  def clear_poses():
      pose = create_transition_pose()
      pose_start = create_transition_pose()
      pose_help = create_transition_pose()
      pose_target = create_transition_pose()
  end

  def do_transition(reference_pose=p[0,0,0,0,0,0], mode=2, keep_rxry=False, a=1.4, v=1.05, r=0.100):
      # the robot will evaluate the current and target workarea
      # after that, the robot will move between the workareas automatically.
      # parameters:
      # reference_pose:   a pose/frame were the robot should work next. If nothing is given, base frame will be used as target
      # keep_rxry:        if true, the robot will keep the orientation of the tool during the movement

      ################# checking #################
      clear_poses()
      workarea_current = check_workarea(get_actual_tcp_pose())    # between 0 and the amount of defined workareas
      workarea_new = check_workarea(reference_pose)               # between 0 and the amount of defined workareas
      reverse_rotation = False

      if (workarea_current != 0 and workarea_new != 0 and workarea_current != workarea_new) or (reference_pose == p[0,0,0,0,0,0]):
          ################# get axisvalues #################
          if (mode == 1):
              pose_start = get_transition_pose_by_workarea(workarea_current)
              pose_target = get_transition_pose_by_workarea(workarea_new)
          elif (mode == 2):
              pose_start = get_transition_pose_by_reference_pose(get_actual_tcp_pose(), RADIUS_TRANSITION_POSES, keep_rxry)
              pose_target = get_transition_pose_by_reference_pose(reference_pose, RADIUS_TRANSITION_POSES, keep_rxry)

          end
          # if (pose_start.crt[1] < 0 and pose_target.crt[1] > 0) or (pose_start.crt[1] > 0 and pose_target.crt[1] < 0):
          #     pose_help = get_transition_pose_by_reference_pose(pose_start.crt, RADIUS_HELPER_POSES)
          # end
          textmsg("Cartesian pose start: ", to_str(pose_start.crt))
          textmsg("Joints pose start: ", to_str(pose_start.jnt))
          textmsg("Qnear pose start: ", to_str(pose_start.q))
          textmsg("Cartesian pose target: ", to_str(pose_target.crt))
          textmsg("Joints pose target: ", to_str(pose_target.jnt))
          textmsg("Qnear pose target: ", to_str(pose_target.q))

          ################# movements #################
          if (pose_help.jnt != [0,0,0,0,0,0]):
              if point_dist(get_actual_tcp_pose(), pose_start.crt) > r and point_dist(pose_start.crt, pose_help.crt) > r:
                  movej(pose_start.jnt, a=a, v=v, r=r)
                  if (point_dist(pose_start.crt, pose_help.crt) > r) and (point_dist(pose_target.crt, pose_help.crt) > r):
                      movej(pose_help.jnt, a=a, v=v, r=r)
                  end
              end
          else:
              if point_dist(get_actual_tcp_pose(), pose_start.crt) > r and point_dist(pose_start.crt, pose_target.crt) > r:
                  movej(pose_start.jnt, a=a, v=v, r=r)
              end
          end
          movej(pose_target.jnt, a=a, v=v)

          ################# checking #################
          workarea_current = check_workarea(get_actual_tcp_pose())    # between 0 and the amount of defined workareas
      else:
          # define error or warning
      end
  end


  # Erläuterung
  # für start wird die aktuelle Position übergeben
  # davon wird die Position für start berechnet. Bei der Orientierung wird entweder nur Rz genommen oder alles bei keep_rxry
  $ 11 "Script: SCRIPT Logs V1.2.script"
  current_state_log = ""
  current_process_log = ""
  current_step_log = ""
  current_warning_log = ""
  current_error_log = ""
  current_hatch_log = ""
  current_centrifuge_log = ""
  current_message_log = "placeholderstring"
  LogLevel=struct(NONE=0, INFO=1, PROCESS=2, WARNING=3, ERROR=4)
  LOGLEVEL=LogLevel.INFO

  def log_message(prefix="", newlog=current_message_log):
      # generates a log message every time its useful
      if (current_message_log != newlog and newlog != ""):
          textmsg(str_cat(prefix, to_str(newlog)))
          current_message_log = to_str(newlog)
      end
  end

  def log_state(newlog):
      # generates a log message every time its useful
      if (current_state_log != newlog and newlog != ""):
          textmsg(str_cat("Machine: ", to_str(newlog)))
          current_state_log = to_str(newlog)
      end
  end

  def log_process(newlog):
      # generates a log message every time its useful
      if (current_process_log != newlog and newlog != ""):
          textmsg(str_cat("Process: ", to_str(newlog)))
          current_process_log = to_str(newlog)
      end
  end

  def log_step(newlog):
      # generates a log message every time its useful
      if (current_step_log != newlog and newlog != ""):
          textmsg(str_cat("Step: ", to_str(newlog)))
          current_step_log = to_str(newlog)
      end
  end

  def log_info(newlog):
      # generates a log message if log level is Info or lower
      if (newlog != "" and LOGLEVEL <= LogLevel.INFO):
          textmsg(str_cat("INFO: ", newlog))
      end
  end

  def log_warning(newlog):
      # generates a log message every time its useful
      if (current_warning_log != newlog and newlog != ""):
          textmsg(str_cat("WARNING: ", to_str(newlog)))
          current_warning_log = to_str(newlog)
      end
  end

  def log_error(newlog):
      # generates a log message every time its useful
      if (current_error_log != newlog and newlog != ""):
          textmsg(str_cat("ERROR: ", to_str(newlog)))
          current_error_log = to_str(newlog)
      end
  end

  def log_hatch_state(newlog):
      # generates a log message every time its useful
      if (current_hatch_log != to_str(newlog) and to_str(newlog) != ""):
          textmsg(str_cat("Hatch_state: ", to_str(newlog)))
          current_hatch_log = to_str(newlog)
      end
  end

  def log_centrifuge_state(newlog):
      # generates a log message every time its useful
      if (current_centrifuge_log != to_str(newlog) and to_str(newlog) != ""):
          textmsg(str_cat("Centrifuge_state: ", to_str(newlog)))
          current_centrifuge_log = to_str(newlog)
      end
  end
  $ 12 "Script: SCRIPT Statistics V1.1.script"
  #*****************************************************
  # customer          :   tbd
  # project name      :   tbd
  #****************************************************
  # controller        :
  # software          :
  #****************************************************
  # author            :   P. Koehnke (+49 1628859904; p.koehnke@unitedrobotics.group)
  # Copyright (c)     :   United Robotics Group Health and Food GmbH
  #                       An der Riede 2
  #                       28816 Stuhr
  #                       Germany
  #****************************************************
  # description       :   statistics script, which tracks the times in different PackML states and let you count objects
  # version:      	:   1.0
  # created           :   20.11.2023
  # updated           :
  #****************************************************
  # modifications     :
  #
  # date              :
  # name              :
  # reason            :
  #****************************************************

  # to save the times persistently, these variables must be defined in the installation file of the robot

  # ===== object counters =====
  def count_up(counters, idx, by):
      counters[idx] = counters[idx] + by
      return counters
  end

  def count_total(counters):
      local i = 0
      local total = 0
      while (i<length(counters)):
          total = total + counters[i]
          i = i + 1
      end
      return total
  end
  # ==========

  # ===== Times =====
  thread Pml_Timer_Thread():
      # STATE_Times is a list of all time values in seconds
      while (True):
          STATE_Times[STATE-1] = STATE_Times[STATE-1] + get_steptime()
          sync()
      end
  end

  thread_timer_handler = run Pml_Timer_Thread()

  def get_time(timer, format="dd/hh/mm/ss"):
      # give the time in seconds
      # the function will return the given time as string in the predefined format
      local days = floor(timer/86400)
      local hours = floor((timer%86400)/3600)
      local minutes = floor((timer%3600)/60)
      local seconds = floor(timer%60)
      return str_cat(str_cat(str_cat(str_cat(str_cat(str_cat(to_str(days), "/"), to_str(hours)), "/"), to_str(minutes)), "/"), to_str(seconds))
  end

  def set_timer(time, format="dd/hh/mm/ss"):
      # give the time as string
      # the function will return the corresponding seconds summed up
      local days_idx = str_find(time, "/", 0)
      local hours_idx = str_find(time, "/", days_idx+1)
      local minutes_idx = str_find(time, "/", hours_idx+1)
      local days = to_num(str_sub(time, 0, days_idx))
      local hours = to_num(str_sub(time, days_idx+1, hours_idx-days_idx-1))
      local minutes = to_num(str_sub(time, hours_idx+1, minutes_idx-hours_idx-1))
      local seconds = to_num(str_sub(time, minutes_idx+1, length(time)-minutes_idx))
      return (days*86400 + hours*3600 + minutes*60 + seconds)
  end
  $ 13 "Script: SCRIPT Vision Config V0.2.script"
  CAM_LM = struct(id=0, type="", size=0, related_itm=0, capture_relation="")
  global CAM_Result = make_list(0, 0, 50)

  def create_landmark(id=0, type="", size=0, related_itm=0, capture_relation=""):
      return struct(id=id, type=type, size=size, related_itm=related_itm, capture_relation=capture_relation)
  end


  CAM_LMs = [
    create_landmark(id=1, type="aruco_7x7", size=0.1, related_itm=1, capture_relation="front_right"),
    create_landmark(id=4, type="aruco_7x7", size=0.1, related_itm=2, capture_relation="straight_left"),
    create_landmark(id=3, type="aruco_7x7", size=0.1, related_itm=2, capture_relation="straight_left"),
    create_landmark(id=8, type="aruco_7x7", size=0.1, related_itm=2, capture_relation="right"),
    create_landmark(id=5, type="aruco_7x7", size=0.1, related_itm=5, capture_relation="left"),
    create_landmark(id=6, type="aruco_7x7", size=0.1, related_itm=2, capture_relation="straight_left")
  ]

  CAM_Capture_Poses = struct(
    front_left = p[0.350,-0.330,0.500,0.353,-0.323,-1.458],
    left = p[0.350,0.000,0.500,0.353,-0.323,-1.458],
    back_left = p[0.350,0.220,0.500,0.353,-0.323,-1.458],
    back_right = p[-0.350,0.000,0.500,0.579,0.240,0.760],
    right = p[-0.350,-0.300,0.500,0.206,0.206,1.561],
    front_right = p[-0.350,-0.400,0.500,0.242,0.903,2.480],
    straight_left = p[0.375,-0.000,0.500,0.815,-0.815,-1.412],
    front = p[0,0,0,0,0,0]
  )

  def get_capture_pose(lm):
      if (lm.capture_relation == "front_left"):
          return CAM_Capture_Poses.front_left
      elif (lm.capture_relation == "left"):
          return CAM_Capture_Poses.left
      elif (lm.capture_relation == "back_left"):
          return CAM_Capture_Poses.back_left
      elif (lm.capture_relation == "back_right"):
          return CAM_Capture_Poses.back_right
      elif (lm.capture_relation == "right"):
          return CAM_Capture_Poses.right
      elif (lm.capture_relation == "straight_left"):
         return CAM_Capture_Poses.straight_left
      else:
          # error
          return get_actual_tcp_pose()
      end
  end
  $ 14 "Script: SCRIPT uLM Factory.script"
  # ############### SCRIPT uLM Factory ##################
  # *****************************************************
  # Customer          :   URG
  # Product Name      :   uLabMobile
  # ****************************************************
  # Controller/Robot  :   UR5e
  # Software          :   URSCRIPT
  # Dependencies      :   Defines Script but mainly independend
  # How To            :   is used by projectconfig to create list of structs full of projectrelated information which are used across the scripts
  # ****************************************************
  # Author            :   D.Kreugel
  # Copyright (c)     :   United Robotics Group Health and Food GmbH
  #                       An der Riede 2
  #                       28816 Stuhr
  #                       Germany
  # ****************************************************
  # Description       :   definition of the datastructures used by the uLM, gives functionality to create a predefined datastructure, is assigned to a global list in projectconfig
  # Version           :   0.2
  # Created           :   18.07.2024
  # Updated           :
  # ****************************************************
  # Modifications     :
  #
  # Date              :
  # Name              :
  # Reason            :
  # ****************************************************
  # TODO              : cleanup useless info and add all other factorys from the other scripts here to have one place to search for such things, documentation

  # DO NOT TOUCH THE DATASTRUCTURES IF YOU DON'T KNOW WHAT YOU DO!
  MAX_ACTIONS=6
  POS_Z=p[0,0,0,0,0,0]
  def create_pattern(id=0, name="", pattern_width=[0, 0], pattern_size=[0, 0], blocked=[-1, -1, -1], direction="X", transpose=False, invert=False, description="default"):
      return struct(
          id = id,
          name = name,
          pattern_width = pattern_width,
          pattern_size = pattern_size,
          blocked = blocked,
          direction = direction,
          transpose = transpose,
          invert = invert,
          description = description
      )
  end

  # item model stores frame related inner and outer patterns
  def create_item_model(inner="", outer="", description="default"):
      return struct(
          inner = inner,
          outer = outer,
          description = description
          )
  end

  # creates a fixed length list cause structs cannot deal with dynamic lists at the moment and an item can have different amount of actions assigned to it
  def create_action_list(values):
      local list = make_list(MAX_ACTIONS, 0, MAX_ACTIONS+1)
      local i = 0
      while (i < values.length()):
          list[i] = values[i]
          i = i + 1
      end
      return list
  end

  def create_item(id=0, ls_item="default", frame=p[0,0,0,0,0,0], actionlist=create_action_list([]), item_model=create_item_model(), lm_id=0, description="default"):
      return struct(
          id = id,
          ls_item = ls_item,
          frame = frame,
          actionlist = create_action_list(actionlist),
          item_model = item_model,
          lm_id = lm_id,
          description = description
      )
  end

  def create_object(id=0, obj_name=0, height=0, width=0, obj_type = 0, description="default"):
      return struct(
          id = id,
          obj_name = obj_name,
          obj_type = obj_type,
          height = height,
          width = width,
          description = description
      )
  end
  # extends object type by sample related information
  def create_sample(obj_id=0, cap_diameter=0, raw_diameter=0, color="", material="", description=""):
      return struct(
      obj_id = obj_id,
      cap_diameter = cap_diameter,
      raw_diameter = raw_diameter,
      color = color,
      material = material,
      description = description)
  end

  # create gripper configs
  def create_gripper_config(gripper_offset=struct(prepick=2, pick=0, place=2), force=0, speed=0, validation=0, object=create_object()):
      gripper_offset.prepick = object.width+gripper_offset.prepick
      gripper_offset.place = object.width+gripper_offset.place
      return struct(
          object = object.obj_name,
          force = force,
          speed = speed,
          validation = validation,
          width = gripper_offset
      )
  end

  def create_manipulator_command(id="", item="", action=0, jig_nbr=-1, obj_nbr=-1, object_type=-1, error_id=0, data=""):
      return struct(
          id = id,
          device = Device.MANIPULATOR,
          item = item,
          action = action,
          jig_nbr = jig_nbr,
          obj_nbr = obj_nbr,
          object_type = object_type,
          error_id = error_id,
          data = data
      )
  end

  def create_amr_command(id="", item="", action=0, target=0, error_id=0, data=""):
      return struct(
          id = id,
          device = Device.AMR,
          item = item,
          action = action,
          target = target,
          error_id = error_id,
          data = data
      )
  end

  def create_camera_command(id="", item="", action=0, attempt=0, error_id=0, data=""):
      return struct(
          id = id,
          device = Device.CAMERA,
          item = item,
          action = action,
          attempt = attempt,
          error_id = error_id,
          data = data
      )
  end

  # Function to create a new  vision struct to assign workspace and skill to an item or a selection
  def create_vision_config(workspace_id="", skill_id="", item_id=-1, target_origin=p[0,0,0,0,0,0], description="default"):
      return struct(
          workspace_id = workspace_id,
          skill_id = skill_id,
          item_id = item_id,
          target_origin = target_origin,
          description = description)
  end

  # extents the vision config by the inspect configuration, this info will be called in the action inspect only
  # item_id is the reference to the item
  # dx is the distance in x direction for one position to the next in the inspection rack
  # dy is the distance in y direction for one position to the next in the inspection rack
  # target origin is the origin coordinate of the first position in the inspectionrack from where the calculation starts
  def create_inspect_config(item_id=0, dx=0, dy=0, target_origin=p[0,0,0,0,0,0], rack_size=[0,0], description="default"):
      return struct(
      item_id = item_id,
      dx = dx,
      dy = dy,
      target_origin = target_origin,
      rack_size = rack_size,
      description = description
      )
  end
   # Function to create a new landmark struct that contains all lm related configurationparameters and will be assigned via item_id
  #def create_landmark(lm_id=0, marker_id=-1, marker_size=0.1, marker_type="aruco_7x7", capture_pos=p[0,0,0,0,0,0], init_frame=p[0,0,0,0,0,0], search_offset=[0,0,0], actual_frame=p[0,0,0,0,0,0], description=""):
    ##  return struct(
     #     lm_id = lm_id,
     #     marker_id = marker_id,
       #   marker_size = marker_size,
    ##      marker_type = marker_type,
    #      capture_pos = capture_pos,
    #      init_frame = init_frame,
    #      search_offset = search_offset,
    #      actual_frame = actual_frame,
  #        description = description)
  #end

  def create_movement(id=0, actionlist=create_action_list([]), hh_approach=POS_Z, h_approach=POS_Z, approach=POS_Z, h_target=POS_Z, target=POS_Z, retract=POS_Z, h_retract=POS_Z, hh_retract=POS_Z, h_frame=POS_Z, frame=POS_Z, speed=1, acceleration=1, description="default"):
  return struct(
      id = id,
      actionlist = actionlist,
      hh_approach = hh_approach,
      h_approach = h_approach,
      approach = approach,
      h_target = h_target,
      target = target,
      retract = retract,
      h_retract = h_retract,
      hh_retract = hh_retract,
      h_frame = h_frame,
      frame = frame,
      speed = speed,
      acceleration = acceleration,
      description = description
  )
  end






  $ 15 "Script: SCRIPT uLM Defines v0.2.script"
  ############# SCRIPT uLM Defines ###############
  #*****************************************************
  # Customer          :   URG
  # Product Name      :   uLabMobile
  #****************************************************
  # Controller/Robot  :   UR5e
  # Software          :   5.17
  # Dependencies      :   Factory Script, Logs Script
  # How To            :   Define Constants depending on the Project, don't go to big in Listsize as it will exceed the URScript limits
  #****************************************************
  # Author            :   D.Kreugel
  # Copyright (c)     :   United Robotics Group Health and Food GmbH
  #                       An der Riede 2
  #                       28816 Stuhr
  #                       Germany
  #****************************************************
  # Description       :   Defines all Enums and Global reachable Varibles/Datastructures
  # Version           :   0.2
  # Created           :   18.07.2024
  # Updated           :
  #****************************************************
  # Modifications     :
  #
  # Date              :
  # Name              :
  # Reason            :
  #****************************************************
  # TODO find better place for the Search Funktions for the Object Lists, documentation


  POS_Z = p[0,0,0,0,0,0]

  # DEFAULTS ROBOT MOVEMENTS
  DEFAULT = struct(SPEED=0.8, ACCELERATION=0.6)

  # ENUMS
  Objects = struct(NONE=0, CC_SAMPLE=1, CC_RACK=2, COAG_SAMPLE=3, COAG_RACK=4, HEMA_SAMPLE=5, HEMA_RACK=6, INPUT_RACK=7, CF_RACK=8, ANY_SAMPLE=9, ANY_RACK=10, TARA_SAMPLE=11, BUTTON=12, XN550_DRAWER=13, COBAS_RACK=14)
  ObjectType = struct(NONE=0,SAMPLE=1,RACK=2, BUTTON=3, DRAWER=4)

  ActionManipulator = struct(NONE=0, PICK=1, PLACE=2, DECAP=12, PUSH=3, RELEASE=21, GRASP=20, MOVE_TO=19, DRAWER_OPEN=51, DRAWER_CLOSE=52)
  ActionAMR = struct(NONE=0, LOAD_MISSION=31, START_MISSION=32, NAVIGATE=33, ACKNOWLEDGE=34, READ=35)
  ActionCamera = struct(NONE=0, INSPECT=16, DETECT=15, DETECT_OBJECTS=17)
  Device = struct(MANIPULATOR=1, AMR=2, CAMERA=3)
  Patterns = struct(NONE="NONE", TARA="TARA", CENTRIFUGE="CENTRIFUGE",CENTRIFUGE_MAGAZINE="CENTRIFUGE_MAGAZINE",SYSMEX_XN550="SYSMEX_XN550",COBAS="COBAS",COBAS_MAGAZINE="COBAS_MAGAZINE",INPUT="INPUT",NOK="NOK",DRAWER_XN550="DRAWER_XN550",ARCHIVE="ARCHIVE")
  CommandStatus = struct(EXECUTED=0, UNFINISHED=1)

  # Constants
  MAX_CAPTURE_ATTEMPTS = 8
  # Maximum Size of the Datastructures
  MAX_ITEM_OBJ = 40
  MAX_GRIPPER_OBJ = 10
  MAX_LANDMARK_OBJ = 10
  MAX_PATTERN_OBJ = 30
  MAX_ITEM_MODEL_OBJ = 20
  MAX_VISION_CONFIG_OBJ = 10
  MAX_CAPTURE_RESULTS = 55
  MAX_MOVEMENT_OBJ = 50

  CON=False

  # for Marburg Approach
  LAST_CAPTURE = make_list(0, "", MAX_CAPTURE_RESULTS)

  # Initialize the Datastructures in order to store related Data and use them in structs without length issues

  OBJECT_MAP = make_list(0 ,create_object(), MAX_ITEM_OBJ)
  ITEM_MAP = make_list(0, create_item(), MAX_ITEM_OBJ)
  ITEM_MODEL_MAP = make_list(0, create_pattern(), MAX_ITEM_MODEL_OBJ)
  GRIPPER_CONFIG_MAP = make_list(0, create_gripper_config(), MAX_PATTERN_OBJ)
  VISION_CONFIG_MAP = make_list(0, create_vision_config(), MAX_VISION_CONFIG_OBJ)
  INSPECT_CONFIG_MAP = make_list(0, create_inspect_config(), MAX_VISION_CONFIG_OBJ)
  LANDMARK_MAP = make_list(0, create_landmark(), MAX_LANDMARK_OBJ)
  MOVEMENT_MAP = make_list(0, create_movement(), MAX_MOVEMENT_OBJ)

  OBJECT_REFERENCE_HEIGHT = 81


  # functions to search in the datastructures which are defined in the factories

  ################# MOVEMENT ###############

  def find_movement_by_frame_and_action(frame,action):
      local i = 0
      local ii = 0
      while (i < MOVEMENT_MAP.length()):
          if (MOVEMENT_MAP[i].frame == frame):
              while(ii < MOVEMENT_MAP[i].actionlist.length()):
                  if (MOVEMENT_MAP[i].actionlist[ii] == action):
                      log_info("Movement found: [" + to_str(MOVEMENT_MAP[i].description) + "]")
                      return MOVEMENT_MAP[i]
                  end
                  ii = ii + 1
              end
              ii = 0
          end
          i = i + 1
      end
      log_warning("no movement found for frame: [" + to_str(frame) + "]")
      return create_movement(frame=frame)  # Return default pattern if not found
  end

  def find_item_by_lsitem_and_action(ls_item, action):
      local i = 0
      while (i < ITEM_MAP.length()):
          if (ITEM_MAP[i].ls_item == ls_item):
              local ii = 0
              while (ii < ITEM_MAP[i].actionlist.length()):
                  if (ITEM_MAP[i].actionlist[ii] == action):
                      log_info("Item found: [" + to_str(ITEM_MAP[i].description) + "]")
                      return ITEM_MAP[i]
                  end
                  ii = ii + 1
              end
          end
          i = i + 1
      end
      log_warning("Item not found for station[" + to_str(ls_item) + "] and action[" + to_str(action) + "]")
      return create_item()  # Return default item if not found
  end
  ################# PATTERN ###################

  def find_pattern_by_name(name):
      local i = 0
      while (i < ITEM_MODEL_MAP.length()):
          if (ITEM_MODEL_MAP[i].name == name):
              log_info("Item Model found: [" + to_str(ITEM_MODEL_MAP[i].description) + "]")
              return ITEM_MODEL_MAP[i]
          end
          i = i + 1
      end
      log_warning("Item Model not found for name[" + to_str(name) + "]")
      return create_pattern()  # Return default pattern if not found
  end

  def is_in_list(list,val):
      local i = 0
      while(i<list.length()):
          if(list[i]==val):
              return True
          end
          i=i+1
      end
      return False
  end

  def get_next_valid_patternslot(item_model, counter):
      local i = 0
      local temp = 0
      local max_slots = item_model.pattern_size[0] * item_model.pattern_size[1]
      log_info("blocked positions:" + to_str(item_model.blocked) + "| current pos: " + to_str(counter))
      while (i < item_model.blocked.length()):
          if(item_model.blocked[i] <= counter and item_model.blocked[i] != -1):
              temp = temp + 1
          end
          i = i + 1
      end

      if(is_in_list(item_model.blocked,counter+temp)):
          while(is_in_list(item_model.blocked,counter+temp)):
              temp=temp+1
          end
      end
      log_info("changed position in rack to nbr:" + to_str(counter+temp))

      return counter+temp

  end

  ################# OBJECT ###################

  # def find_object_by_material(material):
  #   local i = 0
  #   log_info("Trying to find object by color:", to_str(material))
  #   while (i < OBJECT_MAP.length()):
  #       if (OBJECT_MAP[i].material == material):
  #           log_info("Object model found:", to_str(OBJECT_MAP[i]))
  #           return OBJECT_MAP[i]
  #       end
  #       i = i + 1
  #   end
  #   return OBJ_DEFAULT  # Return default pattern if not found
  # end

  def find_object_by_objectname(objectname):
      local i = 0
      #log_info("Trying to find object by color:", to_str(objectname))
      while (i < OBJECT_MAP.length()):
          if (OBJECT_MAP[i].obj_name == objectname):
              log_info("Object Model found: [" + to_str(OBJECT_MAP[i].description) + "]")
              return OBJECT_MAP[i]
          end
          i = i + 1
      end
      log_warning("no Object Model found for objectname:[" + to_str(objectname) + "]")
      return create_object()
  end

  def find_smallest_object():
      local i = 0
      local min_size = OBJECT_MAP[0].height
      #log_info("Trying to find object by color:", to_str(objectname))
      while (i < OBJECT_MAP.length()):
          if (OBJECT_MAP[i].height <= min_size and OBJECT_MAP[i].height != 0):
              log_info("smaller object found: [" + to_str(OBJECT_MAP[i].description) + "]")
              min_size = OBJECT_MAP[i].height
          end
          i = i + 1
      end
      return min_size
  end

  def find_gripper_config_by_objectname(objectname):
  local i = 0
  while (i < GRIPPER_CONFIG_MAP.length()):
      #log_info("gripper config:",to_str(GRIPPER_CONFIG_MAP[i]))
      if (GRIPPER_CONFIG_MAP[i].object == objectname):
          log_info("found gripper parameters [" + to_str(GRIPPER_CONFIG_MAP[i]) + "]")
          return GRIPPER_CONFIG_MAP[i]
      end
      i = i + 1
  end

  log_warning("no gripper parameters found for object type: " + to_str(objectname))
  return create_gripper_config()
  end
  # Function to find a landmark by item
  def find_landmark_by_id(lm_id):
      local i = 0
      while i < LANDMARK_MAP.length():
          if LANDMARK_MAP[i].lm_id == lm_id:
              log_info("found landmark with id(" + to_str(lm_id) + "): [" + to_str(LANDMARK_MAP[i].description) + "]")
              return LANDMARK_MAP[i]
          end
          i = i + 1
      end
      log_warning("landmark not found for lm_id [" + to_str(lm_id) + "]")
      return create_landmark()
  end
  # Function to find a landmark by item
  def find_landmark_by_capture_pos(capture_pos):
      local i = 0
      while i < LANDMARK_MAP.length():
          if LANDMARK_MAP[i].capture_pos == capture_pos:
              log_info("found landmark by capture_pos [" + to_str(LANDMARK_MAP[i].description) + "]")
              return LANDMARK_MAP[i]
          end
          i = i + 1
      end
      log_warning("Landmark not found for capture_pos: [" + to_str(capture_pos) + "]")
      return create_landmark()
  end

  def update_landmark_by_capture_pos(capture_pos, lm_pos):
      local i = 0
      while i < LANDMARK_MAP.length():
          if LANDMARK_MAP[i].capture_pos == capture_pos:
              log_info("updated landmark from [" + to_str(LANDMARK_MAP[i].description) + "]")
              LANDMARK_MAP[i].actual_frame = lm_pos
              return True
          end
          i = i + 1
      end
      log_warning("Landmark not found for capture_pos: [" + to_str(capture_pos) + "]")
      return False
  end

  def update_landmark_by_id(lm_id,lm_pos):
      local i = 0
      while i < LANDMARK_MAP.length():
          if LANDMARK_MAP[i].lm_id == lm_id:
              log_info("updated landmark.actual_frame from [" + to_str(LANDMARK_MAP[i].description + "]"))
              LANDMARK_MAP[i].actual_frame = lm_pos
              return True
          end
          i = i + 1
      end
      log_warning("Landmark not found for lm_id " + to_str(lm_id))
      return False
  end

  def find_vision_config_by_frame(frame):
      local i = 0
      while i < VISION_CONFIG_MAP.length():
          if VISION_CONFIG_MAP[i].capture_pos == frame:
              log_info("Vision Config found: [" + to_str(VISION_CONFIG_MAP[i].description) + "]")
              return VISION_CONFIG_MAP[i]
          end
          i = i + 1
      end
      log_info("Vision Config not found for frame: " + to_str(frame))
      return create_vision_config()
  end

  def find_vision_config_by_itemid(id):
      local i = 0
      while i < VISION_CONFIG_MAP.length():
          if VISION_CONFIG_MAP[i].item_id == id:
              log_info("Vision Config found: [" + to_str(VISION_CONFIG_MAP[i].description) + "]")
              return VISION_CONFIG_MAP[i]
          end
          i = i + 1
      end
      log_info("Vision Config not found for item: " + to_str(id))
      return create_vision_config()
  end

  def find_inspect_config_by_itemid(id):
      local i = 0
      while i < INSPECT_CONFIG_MAP.length():
          if INSPECT_CONFIG_MAP[i].item_id == id:
              log_info("Inspect Config found: [" + to_str(INSPECT_CONFIG_MAP[i].description) + "]")
              return INSPECT_CONFIG_MAP[i]
          end
          i = i + 1
      end
      log_info("Inspect Config not found for item: " + to_str(id))
      return create_inspect_config()
  end
  $ 16 "Script: SCRIPT Device Robotiq Greifer v0.2.script"
  # ############ SCRIPT Device Robotiq Greifer ###############
  # **********************************************************
  # Customer          :   URG
  # Product Name      :   uLabMobile
  # **********************************************************
  # Controller/Robot  :   UR5e
  # Software          :   5.17
  # Dependencies      :   Logs Script, Robotiq Gripper and Gripper Datastructure for args (Factory Script), URCAP Robotiq
  # **********************************************************
  # Author            :   D.Kreugel, P.Köhnke
  # Copyright (c)     :   United Robotics Group Health and Food GmbH
  #                       An der Riede 2
  #                       28816 Stuhr
  #                       Germany
  # *********************************************************
  # Description       :   Gripper Robotiq Device Interface for Robotiq E-Hand Gripper
  # Version           :   0.2
  # Created           :   18.07.2024
  # Updated           :
  # *********************************************************
  # Modifications     :
  #
  # Date              :
  # Name              :
  # Reason            :
  # *********************************************************
  # TODO              :   documentation

  # RobotiQ Gripper
  ROBOTIQ_GRP_CLOSE = 0
  ROBOTIQ_GRP_OPEN = 40

  # #############FORCEMODE###############
  ROBOTIQ_GRP_FORCE = struct(FULL=100, HALF=50, LOW=25, NONE=0)

  # #############SPEED###################
  ROBOTIQ_GRP_SPEED = struct(FAST=100, MEDIUM=50, SLOW=20)

  # ############VALIDATION###############
  ROBOTIQ_GRP_VALIDATION = struct(ON=1, OFF=0, SKIP=-1)

  # struct(prepick=0, pick=0, place=0, force=0, speed=0, validation=0, object_type=0, description="default")
  def gripper_robotiq_activate():
      return rq_activate_and_wait()
  end

  def gripper_robotiq_reset_and_activate():
      return rq_reset_and_activate()
      #return rq_reset()
  end

  def gripper_robotiq_is_activated():
      return rq_is_gripper_activated()
  end

  def gripper_robotiq_get_current_pos_mm():
      return rq_current_pos_mm()
  end
  # Function to check if the RobotiQ gripper has an object
  def gripper_robotiq_has_object():
      result = rq_is_object_detected()
      if result == False:
          log_error("No object detected by the gripper")
      end
      return result
  end

  def gripper_robotiq_move_to_mm(mm):
      if(gripper_robotiq_is_activated() == False):
          gripper_robotiq_activate()
      end
      return rq_move_and_wait_mm(mm)
  end

  def gripper_robotiq_close():
      if(gripper_robotiq_is_activated() == False):
          gripper_robotiq_activate()
      end
      return rq_close_and_wait()
  end

  def gripper_robotiq_open():
      if(gripper_robotiq_is_activated() == False):
          gripper_robotiq_activate()
      end
      return rq_open_and_wait()
  end

  def gripper_robotiq_set_force(force):
      return rq_set_force_norm(force)
  end

  def gripper_robotiq_set_speed(velocity):
      return rq_set_speed_norm(velocity)
  end
  # Function to initialize the RobotiQ gripper
  # args = struct(obj_type = object.obj_type, force = force, speed = speed, validation = validation, width = (prepick=2, pick=0, place=2))
  def gripper_robotiq_init(args):
      log_info("args:"+to_str(args))
      gripper_robotiq_set_force(args.force)
      gripper_robotiq_set_speed(args.speed)
      if(gripper_robotiq_is_activated() == False):
          gripper_robotiq_activate()
      end
      log_info("Robotiq Gripper Initialized with arguments:" + to_str(args))
      return True
  end
  # Function to prepare the RobotiQ gripper for picking
  # args = struct(obj_type = object.obj_type, force = force, speed = speed, validation = validation, width = (prepick=2, pick=0, place=2))
  def gripper_robotiq_prepick(args):
      gripper_robotiq_init(args)

      if(args.width.prepick <= ROBOTIQ_GRP_CLOSE):
          rq_close_and_wait()
      elif(args.width.prepick >= ROBOTIQ_GRP_OPEN):
          rq_open_and_wait()
      else:
          rq_move_and_wait_mm(args.width.prepick)
      end

      log_info("Robotiq Gripper prepick with arguments:" + to_str(args))
      return True
  end

  # Function to place an object using the RobotiQ gripper
  # args = struct(obj_type = object.obj_type, force = force, speed = speed, validation = validation, width = (prepick=2, pick=0, place=2))
  def gripper_robotiq_place(args):
      gripper_robotiq_init(args)

      if(args.width.place <= ROBOTIQ_GRP_CLOSE):
          rq_close_and_wait()
      elif(args.width.place >= ROBOTIQ_GRP_OPEN):
          rq_open_and_wait()
      else:
          rq_move_and_wait_mm(args.width.place)
      end

      log_info("Gripper Place with arguments:"+ to_str(args))
      return True
  end

  # Function to pick an object using the RobotiQ gripper
  # args = struct(obj_type = object.obj_type, force = force, speed = speed, validation = validation, width = (prepick=2, pick=0, place=2))
  def gripper_robotiq_pick(args):
      gripper_robotiq_init(args)

      if(args.width.pick <= ROBOTIQ_GRP_CLOSE):
          rq_close_and_wait()
      elif(args.width.pick >= ROBOTIQ_GRP_OPEN):
          rq_open_and_wait()
      else:
          rq_move_and_wait_mm(args.width.pick)
      end

      log_info("Gripper Pick with arguments:" + to_str(args))

      if args.validation == ROBOTIQ_GRP_VALIDATION.ON:
          if gripper_robotiq_has_object() == False:
              log_error("Validation failed, no object detected")
              return False
          end
      end

      return True
  end


  # def gripper_robotiq_close_and_validate():
  #     rq_close_and_wait()
  #     if gripper_robotiq_has_object() == False:
  #         log_error("Validation failed, no object detected")
  #         return False
  #     else:
  #         return True
  #     end
  # end



  $ 17 "Script: SCRIPT uLM Gripperconfig v0.6.script"
  ############# SCRIPT uLM Gripperconfig ###############
  #*****************************************************
  # Customer          :   URG
  # Product Name      :   uLabMobile
  #****************************************************
  # Controller/Robot  :   UR5e
  # Software          :   UR-Script
  # Dependencies      :   physical Gripper and Datastructure from Factory for args -> Device Script and Implementations of the Functions
  # How To            :   Assign all Functioncalls to the equivalent of the used Device Script
  #****************************************************
  # Author            :   D.Kreugel, P.Köhnke
  # Copyright (c)     :   United Robotics Group Health and Food GmbH
  #                       An der Riede 2
  #                       28816 Stuhr
  #                       Germany
  #****************************************************
  # Description       :   Defines all Gripperm related Parameters and Functions
  # Version           :   0.6
  # Created           :   18.07.2024
  # Updated           :
  #****************************************************
  # Modifications     :   -> at the moment Gripperconfig linked to Robotiq Gripper Device Script
  # Date              :   18.07.2017
  # Name              :   D.Kreugel
  # Reason            :   uLM Standard
  #****************************************************
  # TO DO             : Implement Activate and Reset Routine at the beginning or after an error depending on the state if an Object is gripped or not, documentation



  # GRIPPER DEFINES
  GRIPPER_CLOSE = ROBOTIQ_GRP_CLOSE
  GRIPPER_OPEN = ROBOTIQ_GRP_OPEN
  # #############FORCE###############
  GRIPPER_FORCE = ROBOTIQ_GRP_FORCE
  # #############SPEED###################
  GRIPPER_SPEED = ROBOTIQ_GRP_SPEED
  # ############VALIDATION###############
  GRIPPER_VALIDATION = ROBOTIQ_GRP_VALIDATION

  # takes force in %
  def gripper_set_force(force):
      return gripper_robotiq_set_force(force)
  end

  # takes speed in %
  def gripper_set_speed(velocity):
      return gripper_robotiq_set_speed(velocity)
  end

  def gripper_activate():
      return gripper_robotiq_activate()
  end

  def gripper_reset_and_activate():
      return gripper_robotiq_reset_and_activate()
  end

  def gripper_is_activated():
      return gripper_robotiq_is_activated()
  end

  def gripper_get_current_pos_mm():
      return gripper_robotiq_get_current_pos_mm()
  end

  def gripper_has_object():
      return gripper_robotiq_has_object()
  end

  def gripper_open():
      return gripper_robotiq_open()
  end

  def gripper_close():
      return gripper_robotiq_close()
  end

  def gripper_move_to_pos_mm(mm):
      return gripper_robotiq_move_to_mm(mm)
  end

  # args = struct(obj_type = object.obj_type, force = force, speed = speed, validation = validation, width = (prepick=2, pick=0, place=2))
  def gripper_init(args):
      return gripper_robotiq_init(args)
  end

  # args = struct(obj_type = object.obj_type, force = force, speed = speed, validation = validation, width = (prepick=2, pick=0, place=2))
  def gripper_prepick(args):
      return gripper_robotiq_prepick(args)
  end

  # args = struct(obj_type = object.obj_type, force = force, speed = speed, validation = validation, width = (prepick=2, pick=0, place=2))
  def gripper_pick(args):
      return gripper_robotiq_pick(args)
  end

  # args = struct(obj_type = object.obj_type, force = force, speed = speed, validation = validation, width = (prepick=2, pick=0, place=2))
  def gripper_place(args):
      return gripper_robotiq_place(args)
  end


  # def gripper_close_and_validate():
  #     return gripper_robotiq_close_and_validate()
  # end

  $ 18 "Script: SCRIPT uLM Projectconfig 0.2.script"
  ############# SCRIPT uLM Projectconfig ###############
  #*****************************************************
  # Customer          :   URG
  # Product Name      :   uLabMobile
  #****************************************************
  # Controller/Robot  :   UR5e
  # Software          :   5.17
  # Dependencies      :   Factory Script, Defines Script, relevant project knowledge about objects, patterns, items, commands, vision skills, landmarktypes and movements
  # How To            :   Define Step by Step all Project Data by creating the objects and appending them to the assigned List, if you skip information
  #                       the default value will be assigned -> give as many details as possible as the default values will not work in some cases
  #****************************************************
  # Author            :   D.Kreugel
  # Copyright (c)     :   United Robotics Group Health and Food GmbH
  #                       An der Riede 2
  #                       28816 Stuhr
  #                       Germany
  #****************************************************
  # Description       :   Project Related Configurations -> in the future will be configured by UGO
  # Version           :   0.2
  # Created           :   18.07.2024
  # Updated           :
  #****************************************************
  # Modifications     :
  # Date              :
  # Name              :
  # Reason            :
  #****************************************************
  # TO DO             :  Simplify Rack Assignment, create Enums for Choices that can be made and will be repeated in many projects, documentation

  #

  # Please Import DeviceScripts and Defines Script First as you may wanna use some of the Defined Variables here

  # Define here the Objects that should be handled, add a new Object Type in the defines if necessary
  # create_object(id=0, obj_name=0, height=0, width=0, color="default", material="default", description="default")
  # struct(NONE=0, CC_SAMPLE=1, CC_RACK=2, COAG_SAMPLE=3, COAG_RACK=4, HEMA_SAMPLE=5, HEMA_RACK=6, INPUT_RACK=7, CF_RACK=8, ANY_SAMPLE=9, ANY_RACK=10)
  #create_object(id=0, obj_name=0, height=0, width=0, obj_type = 0, description="default")
  OBJECT_MAP.append(create_object(id=0, obj_name=Objects.NONE, obj_type=ObjectType.NONE, height=0, width=0, description="None Object"))
  OBJECT_MAP.append(create_object(id=1, obj_name=Objects.CC_SAMPLE, obj_type=ObjectType.SAMPLE, height=108, width=15, description="BD Li-Heparin"))
  OBJECT_MAP.append(create_object(id=2, obj_name=Objects.HEMA_SAMPLE, obj_type=ObjectType.SAMPLE, height=81, width=13, description="BD EDTA"))
  OBJECT_MAP.append(create_object(id=3, obj_name=Objects.CC_SAMPLE, obj_type=ObjectType.SAMPLE, height=108, width=15, description="BD Li-Heparin"))
  OBJECT_MAP.append(create_object(id=4, obj_name=Objects.HEMA_SAMPLE, obj_type=ObjectType.SAMPLE, height=81, width=13, description="Sarstedt EDTA"))
  OBJECT_MAP.append(create_object(id=5, obj_name=Objects.CC_SAMPLE, obj_type=ObjectType.SAMPLE, height=110, width=15, description="Sarstedt Serum-Gel"))
  OBJECT_MAP.append(create_object(id=6, obj_name=Objects.ANY_SAMPLE, obj_type=ObjectType.SAMPLE, height=110, width=15, description="Any Sample"))
  OBJECT_MAP.append(create_object(id=7, obj_name=Objects.ANY_RACK, height=150, width=120, description="Any Rack"))
  OBJECT_MAP.append(create_object(id=8, obj_name=Objects.CF_RACK, height=110, width=15, description="Centrifuge Rack"))
  OBJECT_MAP.append(create_object(id=12, obj_name=Objects.COBAS_RACK, height=OBJECT_REFERENCE_HEIGHT, width=20, description="Cobas Rack"))
  OBJECT_MAP.append(create_object(id=9, obj_name=Objects.TARA_SAMPLE, obj_type=ObjectType.SAMPLE, height=110, width=15, description="Tara Sample"))
  OBJECT_MAP.append(create_object(id=10, obj_name=Objects.BUTTON, obj_type=ObjectType.BUTTON, height=0, width=0, description="Button"))
  OBJECT_MAP.append(create_object(id=11, obj_name=Objects.XN550_DRAWER, height=OBJECT_REFERENCE_HEIGHT, width=25, description="XN550 Drawer"))

  #create_sample(obj_id=0, diameter=0, color="", material="", description="")
  SAMPLES = make_list(0,create_sample(),MAX_ITEM_OBJ)
  SAMPLES.append(create_sample(obj_id=1, cap_diameter=17.4, raw_diameter=15.3, color="darkgreen", material="88", description="BD Li-Heparin -> decapped in Cobas"))
  SAMPLES.append(create_sample(obj_id=1, cap_diameter=17.4, raw_diameter=15.3, color="darkgreen", material="80", description="BD Li-Heparin -> decapped in Cobas"))
  SAMPLES.append(create_sample(obj_id=1, cap_diameter=17.4, raw_diameter=15.3, color="darkgreen", material="93", description="BD Li-Heparin -> decapped in archive"))
  SAMPLES.append(create_sample(obj_id=2, cap_diameter=15.5, raw_diameter=12.3, color="violet", material="82", description="BD EDTA -> Sysmex ->Archive"))
  SAMPLES.append(create_sample(obj_id=2, cap_diameter=15.5, raw_diameter=12.3, color="violet", material="91", description="BD EDTA ->Archive"))
  SAMPLES.append(create_sample(obj_id=2, cap_diameter=15.5, raw_diameter=12.3, color="violet", material="96", description="BD EDTA ->Archive"))
  SAMPLES.append(create_sample(obj_id=3, cap_diameter=17.4, raw_diameter=15.3, color="lightgreen", material="88", description="BD Li-Heparin -> decapped in Cobas"))
  SAMPLES.append(create_sample(obj_id=3, cap_diameter=17.4, raw_diameter=15.3, color="lightgreen", material="93", description="BD Li-Heparin -> decapped in Archive"))
  SAMPLES.append(create_sample(obj_id=3, cap_diameter=17.4, raw_diameter=15.3, color="lightgreen", material="97", description="BD Li-Heparin -> decapped in Archive"))
  SAMPLES.append(create_sample(obj_id=4, cap_diameter=15.6, raw_diameter=12.3, color="red", material="82", description="BD EDTA -> Sysmex ->Archive"))
  SAMPLES.append(create_sample(obj_id=4, cap_diameter=15.6, raw_diameter=12.3, color="red", material="91", description="BD EDTA -> Archive"))
  SAMPLES.append(create_sample(obj_id=4, cap_diameter=15.6, raw_diameter=12.3, color="red", material="96", description="BD EDTA -> Archive"))
  SAMPLES.append(create_sample(obj_id=5, cap_diameter=17.4, raw_diameter=15.3, color="brown", material="80", description="Sarstedt Serum-Gel -> decapped in Cobas"))
  SAMPLES.append(create_sample(obj_id=5, cap_diameter=17.4, raw_diameter=15.3, color="brown", material="93", description="Sarstedt Serum-Gel -> decapped in Archive"))

  # Gripper Configurations depending on the Object Type , add new force and speed in the Defines if necessary
  # create_gripper_config(gripper_offset=struct(prepick=2, pick=0, place=2), force=0, speed=0, validation=0, object=create_object())
  GRIPPER_CONFIG_MAP.append(create_gripper_config(gripper_offset=struct(prepick=2, pick=0, place=2), force=GRIPPER_FORCE.HALF, speed=GRIPPER_SPEED.MEDIUM, validation=GRIPPER_VALIDATION.ON, object=find_object_by_objectname(Objects.ANY_SAMPLE)))
  GRIPPER_CONFIG_MAP.append(create_gripper_config(gripper_offset=struct(prepick=2, pick=0, place=2), force=GRIPPER_FORCE.FULL, speed=GRIPPER_SPEED.MEDIUM, validation=GRIPPER_VALIDATION.ON, object=find_object_by_objectname(Objects.ANY_RACK)))
  GRIPPER_CONFIG_MAP.append(create_gripper_config(gripper_offset=struct(prepick=2, pick=0, place=2), force=GRIPPER_FORCE.HALF, speed=GRIPPER_SPEED.MEDIUM, validation=GRIPPER_VALIDATION.ON, object=find_object_by_objectname(Objects.CC_SAMPLE)))
  GRIPPER_CONFIG_MAP.append(create_gripper_config(gripper_offset=struct(prepick=3, pick=0, place=3), force=GRIPPER_FORCE.HALF, speed=GRIPPER_SPEED.MEDIUM, validation=GRIPPER_VALIDATION.ON, object=find_object_by_objectname(Objects.HEMA_SAMPLE)))
  GRIPPER_CONFIG_MAP.append(create_gripper_config(gripper_offset=struct(prepick=4, pick=0, place=4), force=GRIPPER_FORCE.HALF, speed=GRIPPER_SPEED.MEDIUM, validation=GRIPPER_VALIDATION.OFF, object=find_object_by_objectname(Objects.TARA_SAMPLE)))
  GRIPPER_CONFIG_MAP.append(create_gripper_config(gripper_offset=struct(prepick=2, pick=0, place=2), force=GRIPPER_FORCE.FULL, speed=GRIPPER_SPEED.MEDIUM, validation=GRIPPER_VALIDATION.ON, object=find_object_by_objectname(Objects.CF_RACK)))
  GRIPPER_CONFIG_MAP.append(create_gripper_config(gripper_offset=struct(prepick=2, pick=0, place=2), force=GRIPPER_FORCE.FULL, speed=GRIPPER_SPEED.MEDIUM, validation=GRIPPER_VALIDATION.ON, object=find_object_by_objectname(Objects.COBAS_RACK)))
  GRIPPER_CONFIG_MAP.append(create_gripper_config(gripper_offset=struct(prepick=0, pick=0, place=0), force=GRIPPER_FORCE.HALF, speed=GRIPPER_SPEED.MEDIUM, validation=GRIPPER_VALIDATION.OFF, object=find_object_by_objectname(Objects.NONE)))
  GRIPPER_CONFIG_MAP.append(create_gripper_config(gripper_offset=struct(prepick=0, pick=0, place=0), force=GRIPPER_FORCE.HALF, speed=GRIPPER_SPEED.MEDIUM, validation=GRIPPER_VALIDATION.OFF, object=find_object_by_objectname(Objects.BUTTON)))
  GRIPPER_CONFIG_MAP.append(create_gripper_config(gripper_offset=struct(prepick=5, pick=25, place=5), force=GRIPPER_FORCE.HALF, speed=GRIPPER_SPEED.MEDIUM, validation=GRIPPER_VALIDATION.OFF, object=find_object_by_objectname(Objects.XN550_DRAWER)))
  # create Patterns like Racks or Magazines
  # easy if you define x and y regarding to the base coordinate system  if not you have to deal with transpose and or invert
  # create_pattern(id=0, pattern_width=[0, 0], pattern_size=[0, 0], blocked=[-1, -1], obj_name=0, direction="X", transpose=False, invert=False, description="default")
  # Objectss: NONE=0, CC_SAMPLE=1, CC_RACK=2, COAG_SAMPLE=3, COAG_RACK=4, HEMA_SAMPLE=5, HEMA_RACK=6, INPUT_RACK=7, CENTRIFUGE_RACK=8, ANY_SAMPLE=9, ANY_RACK=10
  # ITEM_MODEL_MAP.append(create_pattern(id=0, pattern_width=[0, 0], pattern_size=[0, 0], blocked=[-1, -1, -1],  direction="X", transpose=False, invert=False, description="default"))
  # ITEM_MODEL_MAP.append(create_pattern(id=1, pattern_width=[0.06, 0], pattern_size=[3, 1],  direction="X", description="Tara"))
  # ITEM_MODEL_MAP.append(create_pattern(id=2, pattern_width=[0.183, 0.082], pattern_size=[10, 5], description="Sarstedt 50 D17 Rack"))
  # ITEM_MODEL_MAP.append(create_pattern(id=3, pattern_width=[0.153, 0.067], pattern_size=[10, 5], description="Sarstedt 50 D13 Rack"))
  # ITEM_MODEL_MAP.append(create_pattern(id=4, pattern_width=[0.06, 0.06], pattern_size=[3, 3], blocked=[5, -1, -1], description="Hettich Centrifuge Rack"))
  # ITEM_MODEL_MAP.append(create_pattern(id=5, pattern_width=[0.093, 0.093], pattern_size=[2, 2],  description="Hettich Centrifuge Rack Magazin"))
  # ITEM_MODEL_MAP.append(create_pattern(id=6, pattern_width=[0.08, 0.05], pattern_size=[5, 2], description="Sysmex XN 550 Rack"))
  # ITEM_MODEL_MAP.append(create_pattern(id=7, pattern_width=[0.175, 0.078], pattern_size=[8, 4], description="URG Rack 40 D17"))
  # ITEM_MODEL_MAP.append(create_pattern(id=8, pattern_width=[0.092, 0], pattern_size=[5, 1], description="Cobas Rack"))
  # ITEM_MODEL_MAP.append(create_pattern(id=9, pattern_width=[0.245, 0.123], pattern_size=[3, 5], blocked=[9,11,12], description="Cobas Rack Magazin"))
  # ITEM_MODEL_MAP.append(create_pattern(id=10, pattern_width=[0.237, 0.095], pattern_size=[11, 5], description="Atellica Rack 5x11"))
  # ITEM_MODEL_MAP.append(create_pattern(id=11, pattern_width=[0.237, 0.095], pattern_size=[2, 2], description="Sensors LM"))
  # ITEM_MODEL_MAP.append(create_pattern(id=12, pattern_width=[0.18, 0], pattern_size=[10, 1], description="Sysmex CS2500 Rack"))
  # ITEM_MODEL_MAP.append(create_pattern(id=13, pattern_width=[0.310, 0.075], pattern_size=[13, 4], description="URG RACK 52 - Special Input"))
  # ITEM_MODEL_MAP.append(create_pattern(id=14, pattern_width=[0.075, 0.075], pattern_size=[4, 6], description="URG RACK 24 - Special NoK"))
  # ITEM_MODEL_MAP.append(create_pattern(id=15, pattern_width=[0.120, 0], pattern_size=[2, 1], description="XN550 Drawer"))

  ITEM_MODEL_MAP.append(create_pattern(id=0, name="NONE", pattern_width=[0, 0], pattern_size=[0, 0], blocked=[-1, -1, -1],  direction="X", transpose=False, invert=False, description="default"))
  ITEM_MODEL_MAP.append(create_pattern(id=1, name="TARA", pattern_width=[0.06, 0], pattern_size=[3, 1],  direction="X", description="Tara"))
  ITEM_MODEL_MAP.append(create_pattern(id=4, name="CENTRIFUGE", pattern_width=[0.06, 0.06], pattern_size=[3, 3], blocked=[5, -1, -1], description="Hettich Centrifuge Rack"))
  ITEM_MODEL_MAP.append(create_pattern(id=5, name="CENTRIFUGE_MAGAZINE", pattern_width=[0.093, 0.093], pattern_size=[2, 2],  description="Hettich Centrifuge Rack Magazin"))
  ITEM_MODEL_MAP.append(create_pattern(id=6, name="SYSMEX_XN550", pattern_width=[0.08, 0.05], pattern_size=[5, 2], description="Sysmex XN 550 Rack"))
  ITEM_MODEL_MAP.append(create_pattern(id=8, name="COBAS", pattern_width=[0.092, 0], pattern_size=[5, 1], description="Cobas Rack"))
  ITEM_MODEL_MAP.append(create_pattern(id=9, name="COBAS_MAGAZINE", pattern_width=[0.245, 0.123], pattern_size=[3, 5], blocked=[9,11,12], description="Cobas Rack Magazin"))
  ITEM_MODEL_MAP.append(create_pattern(id=13, name="INPUT", pattern_width=[0.310, 0.075], pattern_size=[13, 4], description="URG RACK 52 - Special Input"))
  ITEM_MODEL_MAP.append(create_pattern(id=14, name="NOK", pattern_width=[0.075, 0.075], pattern_size=[4, 6], description="URG RACK 24 - Special NoK"))
  ITEM_MODEL_MAP.append(create_pattern(id=15, name="DRAWER_XN550", pattern_width=[0.120, 0], pattern_size=[2, 1], description="XN550 Drawer"))
  ITEM_MODEL_MAP.append(create_pattern(id=7, name="ARCHIVE", pattern_width=[0.175, 0.078], pattern_size=[8, 4], description="URG Rack 40 D17"))






  # add a "skill" to the robots skillset the control system will send a string with the ls_item and action and here we will look if we have a matching skill to execute
  # the item_modell defines the patterns which have to be used by the robot on multiple racks and or multiple samples in a rackpattern
  # inner pattern is always dependung on the object that has to be moved and the outer pattern is the pattern for the containers where the objects are stored in.
  # if racks have to be handled it is also an inner pattern cause the object to handle is the rack itself
  # create_item(id=0, ls_item="default", frame=p[0,0,0,0,0,0], actionlist=create_action_list([]), item_model=create_item_model(), lm_id=0, description="default")
  # create_item_model(inner=create_pattern(), outer=create_pattern(), description="default")
  # ITEM_MAP.append(create_item(id=1, ls_item="Home", frame=F1_uLM_Home, actionlist=[ActionManipulator.MOVE_TO], description="uLM Move To Home"))
  # ITEM_MAP.append(create_item(id=2, ls_item="InputStation", frame=F2_uLM_Input, actionlist=[ActionManipulator.PICK, ActionManipulator.PLACE], item_model=create_item_model(inner=Patterns.INPUT), description="uLM Pick and Place samples from Input"))
  # ITEM_MAP.append(create_item(id=3, ls_item="InputCapture", frame=F3_Cap_Input, actionlist=[ActionCamera.INSPECT, ActionManipulator.MOVE_TO], description="uLM Inspect samples from Input and Move To Capture Position"))
  # ITEM_MAP.append(create_item(id=4, ls_item="Bin", frame=F4_uLM_Bin, actionlist=[ActionManipulator.PLACE], description="uLM Place Cap to Bin"))
  # ITEM_MAP.append(create_item(id=5, ls_item="StationaryGripper", frame=F5_uLM_Gripper, actionlist=[ActionManipulator.PICK, ActionManipulator.PLACE, ActionManipulator.DECAP, ActionManipulator.MOVE_TO, ActionManipulator.GRASP, ActionManipulator.RELEASE], description=" uLM stationary gripper"))
  # ITEM_MAP.append(create_item(id=6, ls_item="CobasRack", frame=F6_uLM_Cobas_R, actionlist=[ActionManipulator.PICK, ActionManipulator.PLACE], item_model=create_item_model(outer=Patterns.COBAS_MAGAZINE), description="uLM Cobas Racks Pick and Place"))
  # ITEM_MAP.append(create_item(id=7, ls_item="CobasMagazine", frame=F7_uLM_Coba_Mag, actionlist=[ActionManipulator.PICK, ActionManipulator.PLACE], item_model=create_item_model(inner=Patterns.COBAS, outer=Patterns.COBAS_MAGAZINE), description="uLM Cobas Magazine Samples Pick and Place"))
  # ITEM_MAP.append(create_item(id=8, ls_item="DetectCobasRacks", frame=F8_Cap_Cobas_LM, actionlist=[ActionCamera.DETECT_OBJECTS, ActionManipulator.MOVE_TO], lm_id=2, description="uLM Cobas Rack Detection and Move To Capture"))
  # ITEM_MAP.append(create_item(id=9, ls_item="TaraMagazine", frame=F9_uLM_Tara, actionlist=[ActionManipulator.PICK, ActionManipulator.PLACE], item_model=create_item_model(inner=Patterns.TARA), description="uLM Centrifuge Tara Pick and Place"))
  # ITEM_MAP.append(create_item(id=10, ls_item="CentrifugeCapture", frame=F10_Cap_CF, actionlist=[ActionManipulator.MOVE_TO, ActionCamera.DETECT], lm_id=1, description="Centrifuge Device Move to Capture Pos and Detect Landmarks"))
  # ITEM_MAP.append(create_item(id=11, ls_item="Centrifuge", frame=F11_CF_PiPl, actionlist=[ActionManipulator.PICK, ActionManipulator.PLACE], description="Centrifuge Device Rack Pick and Place"))
  # ITEM_MAP.append(create_item(id=12, ls_item="CentrifugeMagazine", frame=F12_uLM_CF_Mag, actionlist=[ActionManipulator.PICK, ActionManipulator.PLACE], item_model=create_item_model(inner=Patterns.CENTRIFUGE, outer=Patterns.CENTRIFUGE_MAGAZINE), description=" uLM Centrifuge Magazin Pick and Place"))
  # ITEM_MAP.append(create_item(id=13, ls_item="CentrifugeRack", frame=F13_uLM_CF_R, actionlist=[ActionManipulator.PICK, ActionManipulator.PLACE], item_model=create_item_model(outer=Patterns.CENTRIFUGE_MAGAZINE), description="uLM Centrifuge Magazin Pick and Place Racks"))
  # ITEM_MAP.append(create_item(id=14, ls_item="DailyArchive", frame=F14_uLM_Archive, actionlist=[ActionManipulator.PICK, ActionManipulator.PLACE], item_model=create_item_model(inner=Patterns.ARCHIVE), description="uLM Pick and Place samples from Archive Rack"))
  # ITEM_MAP.append(create_item(id=15, ls_item="NokRack", frame=F15_uLM_Nok, actionlist=[ActionManipulator.PICK, ActionManipulator.PLACE], item_model=create_item_model(inner=Patterns.NOK), description="uLM Pick and Place samples from Nok Rack"))
  # ITEM_MAP.append(create_item(id=16, ls_item="CobasInput", frame=F16_Cobas_Input, actionlist=[ActionManipulator.PLACE], description="uLM Place Cobasrack in Cobas Device"))
  # ITEM_MAP.append(create_item(id=17, ls_item="CobasInputCapture", frame=F17_Cobas_Cap, actionlist=[ActionCamera.DETECT, ActionManipulator.MOVE_TO], lm_id=3, description="uLM Place Cobasrack in Cobas Device"))
  # ITEM_MAP.append(create_item(id=18, ls_item="XN550Input", frame=F18_XN550_Input, actionlist=[ActionManipulator.PICK, ActionManipulator.PLACE], item_model=create_item_model(inner=Patterns.SYSMEX_XN550, outer=Patterns.DRAWER_XN550), lm_id=4, description="uLM Pick and Place Samples in or out of XN550 Racks"))
  # ITEM_MAP.append(create_item(id=19, ls_item="XN550Capture", frame=F19_XN550_Cap, actionlist=[ActionCamera.DETECT, ActionManipulator.MOVE_TO], lm_id=4, description="uLM Move To and Capture LM XN550"))
  # ITEM_MAP.append(create_item(id=20, ls_item="XN550Drawer", frame=F20_XN550_Draw, actionlist=[ActionManipulator.DRAWER_OPEN, ActionManipulator.DRAWER_CLOSE], item_model=create_item_model(inner=Patterns.DRAWER_XN550), lm_id=4, description="uLM Open and close Drawer XN550"))
  # ITEM_MAP.append(create_item(id=21, ls_item="XN550Button", frame=F21_XN550_Btn, actionlist=[ActionManipulator.PUSH], lm_id=4, description="uLM Push XN550 Button"))
  # ITEM_MAP.append(create_item(id=22, ls_item="AMR", frame=p[0,0,0,0,0,0], actionlist=[ActionAMR.READ, ActionAMR.LOAD_MISSION, ActionAMR.START_MISSION, ActionAMR.NAVIGATE, ActionAMR.ACKNOWLEDGE], description="all AMR actions"))



  # ITEM_MAP.append(create_item(id=31, ls_item="TestLM", frame=TestLM, actionlist=[ActionManipulator.PICK, ActionManipulator.PLACE], item_model=create_item_model(inner=Rack.SYSMEX_CS2500), lm_id=5, description="LM Test"))
  # Fills the Vision Config List with Projectrelated Data
  # workspaceid and skillid are highly robominds related so probably will not stay like this in the future
  # sample detection: dx and dy are used to calculate the positions in a rack and given by the offset which will be applied in order to assign the sample to a place in the rack
  # create_vision_config(workspace_id="", skill_id="", item_id=-1, capture_pos=p[0,0,0,0,0,0], dx=0, dy=0, target_origin=p[0,0,0,0,0,0], selector="default", description="default")
  # VISION_CONFIG_MAP.append(create_vision_config(workspace_id="96017791-f581-4e9e-93da-6951695fccc8", skill_id="8885cfe1-6784-4293-bd26-52ebdc67bf95", capture_pos=F10_Cap_CF, target_origin=p[0,0,0,0,0,0], item_id=11, description="LM Detect CF"))
  # VISION_CONFIG_MAP.append(create_vision_config(workspace_id="96017791-f581-4e9e-93da-6951695fccc8", skill_id="8885cfe1-6784-4293-bd26-52ebdc67bf95", capture_pos=F8_Cap_Cobas_LM, target_origin=p[0,0,0,0,0,0], item_id=8, description="LM Detect Cobas Racks"))
  # VISION_CONFIG_MAP.append(create_vision_config(workspace_id="8f0ad01c-dc36-4fdd-b295-0b6b4a38b89a", skill_id="afdc9e13-ea83-40d6-a805-bb041453d2e5", capture_pos=F3_Cap_Input, target_origin=F2_uLM_Input, item_id=3, description="Lab Solution Input Capture"))
  # VISION_CONFIG_MAP.append(create_vision_config(workspace_id="96017791-f581-4e9e-93da-6951695fccc8", skill_id="8885cfe1-6784-4293-bd26-52ebdc67bf95", capture_pos=F19_XN550_Cap, target_origin=F18_XN550_Input, item_id=18, description="Input XN550"))
  # VISION_CONFIG_MAP.append(create_vision_config(workspace_id="96017791-f581-4e9e-93da-6951695fccc8", skill_id="8885cfe1-6784-4293-bd26-52ebdc67bf95", capture_pos=F19_XN550_Cap, target_origin=POS_Z, item_id=19, description="LM Detect XN550F"))
  # VISION_CONFIG_MAP.append(create_vision_config(workspace_id="96017791-f581-4e9e-93da-6951695fccc8", skill_id="8885cfe1-6784-4293-bd26-52ebdc67bf95", capture_pos=F10_Cap_CF, target_origin=POS_Z, item_id=10, description="LM Detect CF"))
  # VISION_CONFIG_MAP.append(create_vision_config(workspace_id="96017791-f581-4e9e-93da-6951695fccc8", skill_id="8885cfe1-6784-4293-bd26-52ebdc67bf95", capture_pos=F19_XN550_Cap, target_origin=F20_XN550_Draw, item_id=20, description="Drawer XN550"))
  # VISION_CONFIG_MAP.append(create_vision_config(workspace_id="96017791-f581-4e9e-93da-6951695fccc8", skill_id="8885cfe1-6784-4293-bd26-52ebdc67bf95", capture_pos=F19_XN550_Cap, target_origin=F21_XN550_Btn, item_id=21, description="Button XN550"))
  # VISION_CONFIG_MAP.append(create_vision_config(workspace_id="96017791-f581-4e9e-93da-6951695fccc8", skill_id="8885cfe1-6784-4293-bd26-52ebdc67bf95", capture_pos=TestLMCap, target_origin=p[0,0,0,0,0,0], item_id=30, description="Button XN550"))
  # VISION_CONFIG_MAP.append(create_vision_config(workspace_id="96017791-f581-4e9e-93da-6951695fccc8", skill_id="8885cfe1-6784-4293-bd26-52ebdc67bf95", capture_pos=TestLMCap, target_origin=TestLM, item_id=31, description="Button XN550"))

  # VISION_CONFIG_MAP.append(create_vision_config(workspace_id="96017791-f581-4e9e-93da-6951695fccc8", skill_id="8885cfe1-6784-4293-bd26-52ebdc67bf95", target_origin=p[0,0,0,0,0,0], item_id=11, description="LM Detect CF"))
  # VISION_CONFIG_MAP.append(create_vision_config(workspace_id="96017791-f581-4e9e-93da-6951695fccc8", skill_id="8885cfe1-6784-4293-bd26-52ebdc67bf95", target_origin=p[0,0,0,0,0,0], item_id=8, description="LM Detect Cobas Racks"))
  # VISION_CONFIG_MAP.append(create_vision_config(workspace_id="8f0ad01c-dc36-4fdd-b295-0b6b4a38b89a", skill_id="afdc9e13-ea83-40d6-a805-bb041453d2e5", target_origin=F2_uLM_Input, item_id=3, description="Lab Solution Input Capture"))
  # VISION_CONFIG_MAP.append(create_vision_config(workspace_id="96017791-f581-4e9e-93da-6951695fccc8", skill_id="8885cfe1-6784-4293-bd26-52ebdc67bf95", target_origin=F18_XN550_Input, item_id=18, description="Input XN550"))
  # VISION_CONFIG_MAP.append(create_vision_config(workspace_id="96017791-f581-4e9e-93da-6951695fccc8", skill_id="8885cfe1-6784-4293-bd26-52ebdc67bf95", target_origin=POS_Z, item_id=19, description="LM Detect XN550F"))
  # VISION_CONFIG_MAP.append(create_vision_config(workspace_id="96017791-f581-4e9e-93da-6951695fccc8", skill_id="8885cfe1-6784-4293-bd26-52ebdc67bf95", target_origin=POS_Z, item_id=10, description="LM Detect CF"))
  # VISION_CONFIG_MAP.append(create_vision_config(workspace_id="96017791-f581-4e9e-93da-6951695fccc8", skill_id="8885cfe1-6784-4293-bd26-52ebdc67bf95", target_origin=F20_XN550_Draw, item_id=20, description="Drawer XN550"))
  # VISION_CONFIG_MAP.append(create_vision_config(workspace_id="96017791-f581-4e9e-93da-6951695fccc8", skill_id="8885cfe1-6784-4293-bd26-52ebdc67bf95", target_origin=F21_XN550_Btn, item_id=21, description="Button XN550"))
  # VISION_CONFIG_MAP.append(create_vision_config(workspace_id="96017791-f581-4e9e-93da-6951695fccc8", skill_id="8885cfe1-6784-4293-bd26-52ebdc67bf95", target_origin=p[0,0,0,0,0,0], item_id=30, description="Button XN550"))
  # VISION_CONFIG_MAP.append(create_vision_config(workspace_id="96017791-f581-4e9e-93da-6951695fccc8", skill_id="8885cfe1-6784-4293-bd26-52ebdc67bf95", target_origin=TestLM, item_id=31, description="Button XN550"))

  # local inputrack = find_pattern_by_name("INPUT")
  # INSPECT_CONFIG_MAP.append(create_inspect_config(item_id=3, dx=inputrack.pattern_width[0]/(inputrack.pattern_size[0]-1), dy=inputrack.pattern_width[1]/(inputrack.pattern_size[1]-1), rack_size=inputrack.pattern_size , description="Input Capture"))
  # # Fills the Landmark List with Projectrelated Data
  # # create_landmark(lm_id=0, marker_id=-1, marker_size=0.1, marker_type="aruco_7x7", capture_pos=p[0,0,0,0,0,0], init_frame=p[0,0,0,0,0,0], search_offset=[0,0,0], actual_frame=p[0,0,0,0,0,0], description="")
  # LANDMARK_MAP.append(create_landmark(lm_id=1, marker_id=3, marker_size=0.1, marker_type="aruco_7x7", capture_pos = F10_Cap_CF, init_frame=p[-0.617789, -0.065471, 0.07918, 0.020983, -0.012695, 1.512066], search_offset=[0.15, 0.15, 0.1], actual_frame=p[-0.617789, -0.065471, 0.07918, 0.020983, -0.012695, 1.512066], description="LM CF Lid"))
  # LANDMARK_MAP.append(create_landmark(lm_id=2, marker_id=-1, marker_size=0.0085, marker_type="aruco_4x4", capture_pos = F8_Cap_Cobas_LM, init_frame=p[0,0,0,0,0,0], search_offset=[0.15, 0.15, 0.1], actual_frame=POS_Z, description="LM Cobas Rack Detection"))
  # LANDMARK_MAP.append(create_landmark(lm_id=3, marker_id=0, marker_size=0.1, marker_type="aruco_7x7", capture_pos = F17_Cobas_Cap, init_frame=p[-0.667,-0.194,0.100,0,0,0], search_offset=[0.15, 0.15, 0.1], actual_frame=POS_Z, description="LM Cobas Cap"))
  # LANDMARK_MAP.append(create_landmark(lm_id=4, marker_id=4, marker_size=0.1, marker_type="aruco_7x7", capture_pos = F19_XN550_Cap, init_frame=p[0.124,-0.976,0.355,-0.008,0.025,3.131], search_offset=[0.15, 0.15, 0.1], actual_frame=p[0,0,0,0,0,0], description="LM XN550 Cap"))
  # LANDMARK_MAP.append(create_landmark(lm_id=5, marker_id=0, marker_size=0.1, marker_type="aruco_7x7", capture_pos = TestLMCap, init_frame=p[-0.49,-0.144,0.092,0,-0.008,0.001], search_offset=[0.15, 0.15, 0.1], actual_frame=POS_Z, description="LM Test"))
  # # Configuration of all movement related parameters
  # # create_movement(id=0, hh_approach=POS_Z, h_approach=POS_Z, approach=POS_Z, h_target=POS_Z, target=POS_Z, retract=POS_Z, h_retract=POS_Z, hh_retract=POS_Z, h_frame=POS_Z, frame=POS_Z, speed=1, acceleration=1, description="default")
  # MOVEMENT_MAP.append(create_movement(description="TestLMCap", frame=TestLMCap, actionlist=[ActionManipulator.MOVE_TO]))
  # MOVEMENT_MAP.append(create_movement(description="TestLM", frame=TestLM, actionlist=[ActionManipulator.PICK,ActionManipulator.PLACE],
  #         approach=p[0,0,0.1,0,0,0],
  #         retract=p[0,0,0.1,0,0,0]))
  # MOVEMENT_MAP.append(create_movement(description="Home - MOVE_TO", frame=F1_uLM_Home, actionlist=[ActionManipulator.MOVE_TO]))
  # MOVEMENT_MAP.append(create_movement(description="Input - PICK&PLACE", frame=F2_uLM_Input, actionlist=[ActionManipulator.PICK,ActionManipulator.PLACE],
  #         approach=p[0,0,0.1,0,0,0],
  #         retract=p[0,0,0.1,0,0,0]))
  # MOVEMENT_MAP.append(create_movement(description="Capture Input - MOVE_TO", frame=F3_Cap_Input, actionlist=[ActionManipulator.MOVE_TO]))
  # MOVEMENT_MAP.append(create_movement(description="BIN - PLACE", frame=F4_uLM_Bin, actionlist=[ActionManipulator.PLACE],
  #         approach=p[0,0,0.1,0,0,0],
  #         retract=p[0,0,0.1,0,0,0]))
  # MOVEMENT_MAP.append(create_movement(description="Gripper - Move To", frame=F5_uLM_Gripper, actionlist=[ActionManipulator.MOVE_TO],
  #         approach=p[0,0,0.1,0,0,0]))
  # MOVEMENT_MAP.append(create_movement(description="Gripper - Pick", frame=F5_uLM_Gripper, actionlist=[ActionManipulator.PICK],
  #         retract=p[0,0,0.1,0,0,0]))
  # MOVEMENT_MAP.append(create_movement(description="Gripper - Place", frame=F5_uLM_Gripper, actionlist=[ActionManipulator.PLACE],
  #         approach=p[0,0,0.1,0,0,0]))
  # MOVEMENT_MAP.append(create_movement(description="CobasRack Pick & Place", frame=F6_uLM_Cobas_R, actionlist=[ActionManipulator.PICK,ActionManipulator.PLACE],
  #         approach=p[0,0,0.1,0,0,0],
  #         target=p[0,0,0,0,0,d2r(90)],
  #         retract=p[0,0,0.1,0,0,0]))
  # MOVEMENT_MAP.append(create_movement(description="CobasMagazine Pick & Place", frame=F7_uLM_Coba_Mag, actionlist=[ActionManipulator.PICK,ActionManipulator.PLACE],
  #         approach=p[0,0,0.1,0,0,0],
  #         target=p[0,0,0,0,0,-d2r(90)],
  #         retract=p[0,0,0.1,0,0,0]))
  # MOVEMENT_MAP.append(create_movement(description="Capture Position Cobas Landmarks", frame=F8_Cap_Cobas_LM, actionlist=[ActionManipulator.MOVE_TO]))
  # MOVEMENT_MAP.append(create_movement(description="TaraMagazine - PICK & PLACE", frame=F9_uLM_Tara, actionlist=[ActionManipulator.PICK,ActionManipulator.PLACE],
  #         approach=p[0,0,0.13,0,0,0],
  #         target=p[0,0,0,0,0,-d2r(90)],
  #         retract=p[0,0,0.13,0,0,0]))
  # MOVEMENT_MAP.append(create_movement(description="Capture Position - Centrifuge LM", frame=F10_Cap_CF,actionlist=[ActionManipulator.MOVE_TO]))
  # MOVEMENT_MAP.append(create_movement(description="Pick and Place Racks - Centrifuge Lid", frame=F11_CF_PiPl, actionlist=[ActionManipulator.PICK,ActionManipulator.PLACE],
  #         approach=p[0,0,0.3,0,0,0],
  #         retract=p[0,0,0.3,0,0,0]))
  # MOVEMENT_MAP.append(create_movement(description="Pick and Place Samples - Centrifuge on uLM", frame=F12_uLM_CF_Mag, actionlist=[ActionManipulator.PICK,ActionManipulator.PLACE],
  #         approach=p[0,0,0.13,0,0,0],
  #         retract=p[0,0,0.13,0,0,0]
  #         ))
  # MOVEMENT_MAP.append(create_movement(description="Pick and Place Racks - Centrifuge on uLM", frame=F13_uLM_CF_R, actionlist=[ActionManipulator.PICK,ActionManipulator.PLACE],
  #         approach=p[0,0,0.15,0,0,0],
  #         retract=p[0,0,0.15,0,0,0]
  #         ))

  # MOVEMENT_MAP.append(create_movement(description="Pick and Place Samples XN550 Racks in Device", frame=F18_XN550_Input, actionlist=[ActionManipulator.PICK,ActionManipulator.PLACE],
  #         approach=p[0,0,0.1,0,0,0],
  #         target = p[0,0,0,0,0,d2r(90)],
  #         retract=p[0,0,0.1,0,0,0]
  #         ))
  # MOVEMENT_MAP.append(create_movement(description="Capture LM XN550", frame=F19_XN550_Cap, actionlist=[ActionManipulator.MOVE_TO]))
  # MOVEMENT_MAP.append(create_movement(description="Open XN550 Drawer ", frame=F20_XN550_Draw, actionlist=[ActionManipulator.DRAWER_OPEN],
  #         h_approach=p[0.07,0,0.1,0,0,0],
  #         approach=p[0,0,0.1,0,0,0],
  #         target = p[0,0,0,0,0,d2r(90)],
  #         retract=p[0.07,0,0,0,0,0],
  #         h_retract=p[0.07,0,0.1,0,0,0]
  #         ))
  # MOVEMENT_MAP.append(create_movement(description="Close XN550 Drawer ", frame=F20_XN550_Draw, actionlist=[ActionManipulator.DRAWER_CLOSE],
  #         h_approach=p[0.07,0,0.1,0,0,0],
  #         approach=p[0.07,0,0,0,0,0],
  #         target = p[0,0,0,0,0,d2r(90)],
  #         retract=p[0,0,0.1,0,0,0],
  #         h_retract=p[0.07,0,0.1,0,0,0]
  #         ))
  # MOVEMENT_MAP.append(create_movement(description="Push XN550 Button ", frame=F21_XN550_Btn, actionlist=[ActionManipulator.PUSH],
  #         approach=p[0,0,0.15,0,0,0],
  #         retract=p[0,0,0.15,0,0,0]
  #         ))
  # MOVEMENT_MAP.append(create_movement(description="Capture Position 2 Input", frame=F_Cap_Input2,actionlist=[ActionManipulator.MOVE_TO]))



  $ 19 "Script: SCRIPT Objects V0.1.script"
  #*****************************************************
  # customer          :   INTERNAL
  # project name      :
  #****************************************************
  # controller        :   UR
  # software          :   5.17.3
  #****************************************************
  # author            :   P. Koehnke
  # Copyright (c)     :   United Robotics Group
  #                       An der Riede 2
  #                       28816 Stuhr
  #                       Germany
  #****************************************************
  # description       :   object database
  # version:      	:   0.1
  # created           :   09.10.2024
  # updated           :
  #****************************************************
  # modifications     :
  #
  # date              :
  # name              :
  # reason            :
  #****************************************************

  def create_object_2(id=0, name="", type=0, dimension=struct(length=0, width=0, height=0, diameter=0), gripper_offset=p[0,0,0,0,0,0]):
      return struct(id=id, name=name, type=type, dimension=dimension, gripper_offset=gripper_offset)
  end

  OBJ = create_object_2()
  OBJs = make_list(0, create_object_2(), 50)

  OBJs.append(create_object_2(id=1, name="rack centrifuge", type=1, dimension=struct(length=0, width=0, height=0.106, diameter=0.020), gripper_offset=p[0,0,0.095,0,0,2.356]))
  OBJs.append(create_object_2(id=2, name="sample tube 1", type=2, dimension=struct(length=0, width=0, height=0.106, diameter=0.015), gripper_offset=p[0,0,0,0,0,0]))
  OBJs.append(create_object_2(id=3, name="rack sarstedt", type=3, dimension=struct(length=0, width=0, height=0.100, diameter=0.020), gripper_offset=p[0,0,0,0,0,0]))
  OBJs.append(create_object_2(id=4, name="Lab bottle", type=4, dimension=struct(length=0, width=0, height=0.100, diameter=0.030), gripper_offset=p[0,0,0.2,0,0,0]))
  OBJs.append(create_object_2(id=5, name="Vial", type=5, dimension=struct(length=0, width=0, height=0.100, diameter=0.0275), gripper_offset=p[0,0,0,0,0,0]))
  OBJs.append(create_object_2(id=6, name="Container_S", type=6, dimension=struct(length=0.09, width=0.09, height=0.185, diameter=0.080), gripper_offset=p[0,0,0,0,0,0]))
  OBJs.append(create_object_2(id=7, name="Target_container", type=7, dimension=struct(length=0.06, width=0.06, height=0.134, diameter=0.05), gripper_offset=p[0,0,0,0,0,0]))
  OBJs.append(create_object_2(id=8, name="Spatula", type=8, dimension=struct(length=0.03, width=0.03, height=0.23, diameter=0.05), gripper_offset=p[0,0,0,0,0,0]))

  def create_jig_2(id=0, name="", type=0, capacity=0, jig_offset=p[0,0,0,0,0,0]):
      # iformation about used jigs
      return struct(id=id, name=name, type=type, capacity=capacity, jig_offset=jig_offset)
  end

  JIG2 = create_jig_2()
  JIGs = make_list(0, create_jig_2(), 20)

  JIGs.append(create_jig_2(id=1, name="3FG", type=1, capacity=1, jig_offset=p[0,0,0,0,0,0]))
  JIGs.append(create_jig_2(id=2, name="jig input", type=2, capacity=1, jig_offset=p[0,0,0,0,0,-3.927]))
  JIGs.append(create_jig_2(id=3, name="jig output", type=3, capacity=1, jig_offset=p[0,0,0,0,0,0.78]))
  JIGs.append(create_jig_2(id=6, name="jig bin", type=6, capacity=1, jig_offset=p[0,0,0,0,0,0]))
  JIGs.append(create_jig_2(id=7, name="jig sarstedt racks", type=7, capacity=1, jig_offset=p[0,0,-0.02,0,0,0]))
  JIGs.append(create_jig_2(id=8, name="NoK Bin", type=8, capacity=1, jig_offset=p[0,0,0,0,0,0]))
  JIGs.append(create_jig_2(id=9, name="Pick bott jig", type=9, capacity=1, jig_offset=p[0,0,0,0,0,0]))
  JIGs.append(create_jig_2(id=10, name="Place bott jig", type=10, capacity=1, jig_offset=p[0,0,0,0,0,0]))
  JIGs.append(create_jig_2(id=11, name="bottle shake jig", type=11, capacity=1, jig_offset=p[0,0,0,0,0,0]))
  JIGs.append(create_jig_2(id=12, name="Pick Vial jig", type=12, capacity=1, jig_offset=p[0,0,0,0,0,0]))
  JIGs.append(create_jig_2(id=13, name="Place Vial jig", type=13, capacity=1, jig_offset=p[0,0,0,0,0,0]))
  JIGs.append(create_jig_2(id=14, name="Liquid transfer jig", type=14, capacity=1, jig_offset=p[0,0,0,0,0,0]))
  JIGs.append(create_jig_2(id=15, name="Pick station jig", type=15, capacity=1, jig_offset=p[0,0,0,0,0,0]))
  JIGs.append(create_jig_2(id=16, name="Place station jig", type=16, capacity=1, jig_offset=p[0,0,0,0,0,0]))
  $ 20 "Script: krish.script"
  def dynamic_upward_motion(distance,duration):
  	speed=distance/duration
  	speed_vector = [0, 0, speed, 0, 0, 0]
  	time_elapsed = 0
  	time_step = 1
  	while time_elapsed < duration:
  		speedl(speed_vector, 0.1, time_step)
  		sleep(time_step)
  		time_elapsed = time_elapsed + time_step
  	end
  	stopl(0.5)
  end
  dynamic_upward_motion(distance, duration)


  def get_weight():
  	socket_open("192.168.12.190", 3002)
  	textmsg("socket opened successfully!")
  	socket_send_string("GET_WEIGHT")
  	sync()
  	sleep(0.5)
  	receiveFromServ = socket_read_ascii_float(6)
  	while (receiveFromServ[0] <1):
  		sleep(0.5)
  		receiveFromServ = socket_read_ascii_float(1)
  		textmsg("retrying read:", receiveFromServ)
  	end
  	textmsg("Received weight:", receiveFromServ[1])
  	socket_close()
  	return receiveFromServ[1]
  end

  get_weight()
  $ 21 "BeforeStarts"
  $ 22 "uLM"
  $ 23 "CMD_Stop≔ False "
  global CMD_Stop=  False
  $ 24 "CMD_Abort≔ False "
  global CMD_Abort=  False
  $ 25 "CMD_Clear≔ False "
  global CMD_Clear=  False
  $ 26 "STATE≔1"
  global STATE=1
  $ 27 "STATE_Info≔''"
  global STATE_Info=""
  $ 28 "ARM_Referenced≔ False "
  global ARM_Referenced=  False
  $ 29 "zero_ftsensor()"
  zero_ftsensor()
  $ 30 "poses init"
  $ 31 "PSE_A≔p[0,0,0,0,0,0]"
  global PSE_A=p[0,0,0,0,0,0]
  $ 32 "PSE_A_H≔p[0,0,0,0,0,0]"
  global PSE_A_H=p[0,0,0,0,0,0]
  $ 33 "PSE_R≔p[0,0,0,0,0,0]"
  global PSE_R=p[0,0,0,0,0,0]
  $ 34 "PSE_R_H≔p[0,0,0,0,0,0]"
  global PSE_R_H=p[0,0,0,0,0,0]
  $ 35 "PSE_T≔p[0,0,0,0,0,0]"
  global PSE_T=p[0,0,0,0,0,0]
  $ 36 "PSE_T_H≔p[0,0,0,0,0,0]"
  global PSE_T_H=p[0,0,0,0,0,0]
  $ 37 "PSE_C_E≔p[0,0,0,0,0,0]"
  global PSE_C_E=p[0,0,0,0,0,0]
  $ 38 "PSE_C_H≔p[0,0,0,0,0,0]"
  global PSE_C_H=p[0,0,0,0,0,0]
  $ 39 "PSE_C_S≔p[0,0,0,0,0,0]"
  global PSE_C_S=p[0,0,0,0,0,0]
  $ 40 "init_home_by_cartesian_pose(p[0,-0.400,0.300,0,0,0])"
  init_home_by_cartesian_pose(p[0,-0.400,0.300,0,0,0])
  $ 41 "Clearing"
  $ 42 "reset_error()"
  reset_error()
  $ 43 "reset_warning()"
  reset_warning()
  $ 44 "uGo"
  $ 46 "ugo_init( True ,'http://192.168.12.120:10001')"
  ugo_init(  True  ,"http://192.168.12.120:10001")
  $ 47 "ugo_update_outputs()"
  ugo_update_outputs()
  $ 48 "App"
  $ 49 "'ADD APPLICATION SPECIFIC COMMANDS'"
  # 'ADD APPLICATION SPECIFIC COMMANDS'
  $ 50 "Tools"
  $ 51 "OBJ_Picked≔gripper_has_object()"
  global OBJ_Picked=gripper_has_object()
  $ 52 "If OBJ_Picked"
  if (OBJ_Picked):
    # begin: URCap Program Node
    #   Source: Robotiq_Grippers, 1.8.4.4844, Robotiq Inc.
    #   Type: Gripper Activate
    $ 53 "Gripper Activate"

    kill rq_gripper_communication_thread
    rq_gripper_communication_thread_started = False

    rq_init_comm_if_connected(9, "1")
    rq_init_comm_if_connected(2, "2")
    rq_init_comm_if_connected(3, "3")
    rq_init_comm_if_connected(4, "4")
    rq_print_connected_grippers()
    rq_gripper_communication_thread = run rq_gripper_communication()

    while(not rq_gripper_communication_thread_started):
        sync()
    end

    rq_set_max_current_for_all_grippers()

    reset_and_activate = False

    rq_activate_all_grippers(False)
    # end: URCap Program Node
  else:
    $ 54 "Else" "noBreak"
    # begin: URCap Program Node
    #   Source: Robotiq_Grippers, 1.8.4.4844, Robotiq Inc.
    #   Type: Gripper Activate
    $ 55 "Gripper Reset and Activate"

    kill rq_gripper_communication_thread
    rq_gripper_communication_thread_started = False

    rq_init_comm_if_connected(9, "1")
    rq_init_comm_if_connected(2, "2")
    rq_init_comm_if_connected(3, "3")
    rq_init_comm_if_connected(4, "4")
    rq_print_connected_grippers()
    rq_gripper_communication_thread = run rq_gripper_communication()

    while(not rq_gripper_communication_thread_started):
        sync()
    end

    rq_set_max_current_for_all_grippers()

    reset_and_activate = True

